// TIA Portal V21 export
// export: Created 2026-11-10T07:35:24.5270971Z, ExportSetting WithDefaults, DisplayName Totally Integrated Automation Portal, DisplayVersion V21 Update 3, DisplayName STEP 7 Professional, DisplayVersion V21 Update 3, DisplayName STEP 7 Safety, DisplayVersion V21, DisplayName Tech WebApplication, DisplayVersion V21, DisplayName WinCC Basic/Comfort/Advanced, DisplayVersion V21 Update 3, DisplayName WinCC Unified, DisplayVersion V21 Update 3
FUNCTION_BLOCK "FB_Lad_ex161"   // FB62, LAD
{ S7_Optimized_Access := 'TRUE' }
VERSION : 0.1
// stored: AutoNumber true, IsIECCheckEnabled false, IsRetainMemResEnabled false, MemoryReserve 100, SetENOAutomatically false, UDAEnableTagReadback false
   VAR_INPUT
      v_ioid : Byte;
      v_laddr : HW_MODULE;
      v_ret_val : Int;
   END_VAR
   VAR_OUTPUT
      v_area : Byte;
      v_rack : Word;
      v_slot : Word;
      v_subaddr : Word;
   END_VAR
BEGIN

REGION Network 1: LGC_GADR - Determine slot from hardware identifier
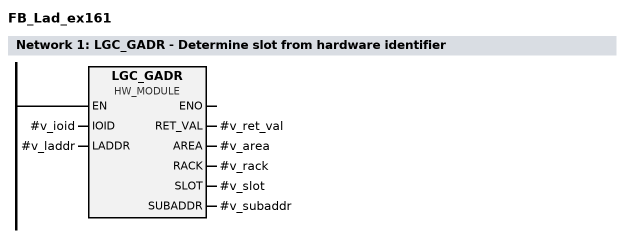
   RUNG wire#powerrail
      { S7_Templates := "laddr_type := HW_MODULE" } LGC_GADR(IOID := #v_ioid, LADDR := #v_laddr, RET_VAL => #v_ret_val, AREA => #v_area, RACK => #v_rack, SLOT => #v_slot, SUBADDR => #v_subaddr)
   END_RUNG
   // the same network as SCL:
   #v_ret_val := LGC_GADR(IOID := #v_ioid,
                          LADDR := #v_laddr,
                          AREA => #v_area,
                          RACK => #v_rack,
                          SLOT => #v_slot,
                          SUBADDR => #v_subaddr);
END_REGION
END_FUNCTION_BLOCK
